// Ab Z1-Position fZ1_mm gilt der Vorschub fFeed_mm_s.
{attribute 'pack_mode' := '1'}
TYPE ST_FeedPoint :
STRUCT
    fZ1_mm : LREAL;
    fFeed_mm_s : LREAL;
END_STRUCT
END_TYPE

(* stored: Version 1.1.0.1
   DUT ST_FeedPoint: Id {9edd77d3-96c3-5ce6-a1b6-20f749bfba40} *)
